// TIA Portal V18 export
TYPE "UDT_DadosEquipScala"
   STRUCT
      Bool0 : Bool;
      Bool1 : Bool;
      Bool2 : Bool;
      Bool3 : Bool;
      Bool4 : Bool;
      Bool5 : Bool;
      Bool6 : Bool;
      Bool7 : Bool;
      Bool8 : Bool;
      Bool9 : Bool;
      Bool10 : Bool;
      Bool11 : Bool;
      Bool12 : Bool;
      Bool13 : Bool;
      Bool14 : Bool;
      Bool15 : Bool;
   END_STRUCT;
END_TYPE
